// TIA Portal V18 export
TYPE "InterlockMdz_in"
   STRUCT
      StationInterlock_APLC_Input : Array[1.."Station_Setup_Const"] of Struct
         PositionInterlock_APLC_Input : Array[1.."Position_Setup_Const"] of Struct
            LoginInterlock_APLC : Bool;
            EquipmentInterlock_APLC_Input : Array[1.."Equipment_Setup_Const"] of Struct
               SignalInterlock_APLC_Input : Array[1.."Signal_Setup_Const"] of Bool;
            END_STRUCT;
         END_STRUCT;
      END_STRUCT;
   END_STRUCT;
END_TYPE
